(* IEC 61131-3 sources: plcassist-cli/packages/volt-lsp-iec/test-corpus/bakon-nano/Device/Plc Logic/Application/POUs/Calculations (part 4) *)

(* ---- Calc_BottomPos.prg ---- *)
PROGRAM Calc_BottomPos
VAR
END_VAR

//Bereken diepste positie van Z-as (Hoogste) afhankelijk van geselecteerd product plaat.

CASE g_HMI_RCP_Parameters.nProductType  OF
	Prod_Tray_Rectangle_1x1:
		g_sCalculated.rBottomZPos		:= g_HMI_MCH_Parameters.rBottomZPosTrayLarge - g_HMI_RCP_Parameters.rStopHeightKnife;
		g_sCalculated.rAboveProductPos	:= MIN((g_HMI_MCH_Parameters.rBottomZPosTrayLarge - g_HMI_RCP_Parameters.rStartHeightKnife - C_rExtraMarginKnifeHeight),(g_HMI_MCH_Parameters.rBottomZPosTrayLarge - g_HMI_MCH_Parameters.rProdHeightTrayMinimum));
		g_sCalculated.rCrashCheckHeight	:= (g_HMI_MCH_Parameters.rBottomZPosTrayLarge - g_HMI_MCH_Parameters.rProdHeightTrayMinimum + 8); // + 5mm
	Prod_Tray_Rectangle_1x2:
		g_sCalculated.rBottomZPos	:= g_HMI_MCH_Parameters.rBottomZPosTraySmall - g_HMI_RCP_Parameters.rStopHeightKnife;
		g_sCalculated.rAboveProductPos := MIN((g_HMI_MCH_Parameters.rBottomZPosTraySmall - g_HMI_RCP_Parameters.rStartHeightKnife - C_rExtraMarginKnifeHeight),(g_HMI_MCH_Parameters.rBottomZPosTraySmall - g_HMI_MCH_Parameters.rProdHeightTrayMinimum));
		g_sCalculated.rCrashCheckHeight	:= (g_HMI_MCH_Parameters.rBottomZPosTraySmall - g_HMI_MCH_Parameters.rProdHeightTrayMinimum + 8); // + 5mm
	Prod_Tray_Rectangle_2x1:		(* V07.01 *)
		g_sCalculated.rBottomZPos		 := g_HMI_MCH_Parameters.rBottomZPosTrayDouble - g_HMI_RCP_Parameters.rStopHeightKnife;
		g_sCalculated.rAboveProductPos := MIN((g_HMI_MCH_Parameters.rBottomZPosTrayDouble - g_HMI_RCP_Parameters.rStartHeightKnife - C_rExtraMarginKnifeHeight),(g_HMI_MCH_Parameters.rBottomZPosTrayDouble - g_HMI_MCH_Parameters.rProdHeightTrayMinimum));
		g_sCalculated.rCrashCheckHeight	:= (g_HMI_MCH_Parameters.rBottomZPosTrayDouble - g_HMI_MCH_Parameters.rProdHeightTrayMinimum + 8); // + 5mm
	Prod_Tray_Rectangle_1x4:
		g_sCalculated.rBottomZPos	:= g_HMI_MCH_Parameters.rBottomZPosTrayTriple - g_HMI_RCP_Parameters.rStopHeightKnife;
		g_sCalculated.rAboveProductPos := MIN((g_HMI_MCH_Parameters.rBottomZPosTrayTriple - g_HMI_RCP_Parameters.rStartHeightKnife - C_rExtraMarginKnifeHeight),(g_HMI_MCH_Parameters.rBottomZPosTrayTriple - g_HMI_MCH_Parameters.rProdHeightTrayMinimum));
		g_sCalculated.rCrashCheckHeight	:= (g_HMI_MCH_Parameters.rBottomZPosTrayTriple -g_HMI_MCH_Parameters.rProdHeightTrayMinimum + 8); // + 5mm
	Prod_Round_POC_2x1:
		g_sCalculated.rBottomZPos	:= g_HMI_MCH_Parameters.rBottomZPosRound - g_HMI_RCP_Parameters.rStopHeightKnife;
		g_sCalculated.rAboveProductPos := MIN((g_HMI_MCH_Parameters.rBottomZPosRound - g_HMI_RCP_Parameters.rStartHeightKnife - C_rExtraMarginKnifeHeight),(g_HMI_MCH_Parameters.rBottomZPosRound - 10));	(* altijd minimaal 10 mm *)
		g_sCalculated.rCrashCheckHeight	:= (g_HMI_MCH_Parameters.rBottomZPosRound - g_HMI_MCH_Parameters.rProdHeightTrayMinimum + 8); // + 5mm
	Prod_Round_POC_2x2:
		g_sCalculated.rBottomZPos	:= g_HMI_MCH_Parameters.rBottomZPosRoundQuatro - g_HMI_RCP_Parameters.rStopHeightKnife;
		g_sCalculated.rAboveProductPos := MIN((g_HMI_MCH_Parameters.rBottomZPosRoundQuatro - g_HMI_RCP_Parameters.rStartHeightKnife - C_rExtraMarginKnifeHeight),(g_HMI_MCH_Parameters.rBottomZPosRoundQuatro - 10));	(* altijd minimaal 10 mm *)
		g_sCalculated.rCrashCheckHeight	:= (g_HMI_MCH_Parameters.rBottomZPosRoundQuatro - g_HMI_MCH_Parameters.rProdHeightTrayMinimum + 8); // + 5mm
	Prod_Slab_Rectangle_2x1:
		g_sCalculated.rBottomZPos	:= g_HMI_MCH_Parameters.rBottomZPosSlabDouble - g_HMI_RCP_Parameters.rStopHeightKnife;
		g_sCalculated.rAboveProductPos := MIN((g_HMI_MCH_Parameters.rBottomZPosSlabDouble - g_HMI_RCP_Parameters.rStartHeightKnife - C_rExtraMarginKnifeHeight),(g_HMI_MCH_Parameters.rBottomZPosSlab - 10));
		g_sCalculated.rCrashCheckHeight	:= (g_HMI_MCH_Parameters.rBottomZPosSlabDouble - g_HMI_MCH_Parameters.rProdHeightTrayMinimum + 8); // + 5mm
ELSE
		g_sCalculated.rBottomZPos	:= g_HMI_MCH_Parameters.rBottomZPosSlab - g_HMI_RCP_Parameters.rStopHeightKnife;
		g_sCalculated.rAboveProductPos := MIN((g_HMI_MCH_Parameters.rBottomZPosSlab - g_HMI_RCP_Parameters.rStartHeightKnife - C_rExtraMarginKnifeHeight),(g_HMI_MCH_Parameters.rBottomZPosSlab - 10));
		g_sCalculated.rCrashCheckHeight	:= (g_HMI_MCH_Parameters.rBottomZPosSlab - g_HMI_MCH_Parameters.rProdHeightTrayMinimum + 8); // + 5mm
END_CASE

g_sCalculated.rCrashCheckHeight := MIN(g_sCalculated.rCrashCheckHeight, g_sCalculated.rBottomZPos-1);

IF g_HMI_MachCommand.bScanMode THEN
		g_sCalculated.rBottomZPos	:= MIN(g_HMI_MCH_Parameters.rBottomZPosSlab,
										MIN(g_HMI_MCH_Parameters.rBottomZPosSlabDouble,
										MIN(g_HMI_MCH_Parameters.rBottomZPosRoundQuatro,
										MIN(g_HMI_MCH_Parameters.rBottomZPosRound,
										MIN(g_HMI_MCH_Parameters.rBottomZPosTrayDouble,
										MIN(g_HMI_MCH_Parameters.rBottomZPosTrayLarge,
										MIN(g_HMI_MCH_Parameters.rBottomZPosTraySmall,
										g_HMI_MCH_Parameters.rBottomZPosTrayTriple)))))));
		g_sCalculated.rAboveProductPos := 0;
END_IF

g_sCalculated.rAboveProductPos := SEL(g_sMACH.MCL.bActCleaning,g_sCalculated.rAboveProductPos,0); //AC Correctie voor schoonmaak bedrijf waarbij er nog geen bottompos is ingesteld

END_PROGRAM

(* ---- Calc_Init.prg ---- *)
PROGRAM Calc_Init
VAR
	Cnt_pos: INT;
END_VAR

(* Init array *)
FOR Cnt_pos := 1 TO (C_wNumberOfMotionObjects -1)  BY 1 DO
	g_aCuttingPositions[Cnt_pos].X_Target			:=-50;
	g_aCuttingPositions[Cnt_pos].Y_Target			:=-50;
	g_aCuttingPositions[Cnt_pos].A_Target			:=-50;
	g_aCuttingPositions[Cnt_pos].K_Target			:= 0;
	g_aCuttingPositions[Cnt_pos].bPushAwayProduct 	:= FALSE;
	g_aCuttingPositions[Cnt_pos].rPushAwayDistance 	:= 0;
	g_aCuttingPositions[Cnt_pos].bCutPosPossible 	:= TRUE;
	g_aCuttingPositions[Cnt_pos].bCrashDetectCheck 	:= FALSE;
END_FOR

FOR Cnt_pos := 1 TO 100 BY 1 DO
	g_aWastePositions[Cnt_pos].X_Target				:=-50;
	g_aWastePositions[Cnt_pos].Y_Target				:=-50;
	g_aWastePositions[Cnt_pos].A_Target				:=-50;
	g_aWastePositions[Cnt_pos].K_Target				:= 0;
	g_aWastePositions[Cnt_pos].bPushAwayProduct 	:= FALSE;
	g_aWastePositions[Cnt_pos].rPushAwayDistance 	:= 0;
	g_aWastePositions[Cnt_pos].bCutPosPossible 		:= TRUE;
	g_aWastePositions[Cnt_pos].bCrashDetectCheck	:= FALSE;
END_FOR

(*Minimale Afvalrand limieten bepalen*)
CASE G_HMI_RCP_Parameters.nProductType OF
	Prod_Tray_Rectangle_1x2, Prod_Tray_Rectangle_1x1, Prod_Tray_Rectangle_1x4, Prod_Tray_Rectangle_2x1 :	(* Tray products *)
	g_HMI_RCP_Parameters.rSizeTrimRight := MAX( g_HMI_RCP_Parameters.rSizeTrimRight, 0);
	g_HMI_RCP_Parameters.rSizeTrimLeft 	:= MAX( g_HMI_RCP_Parameters.rSizeTrimLeft, 0);
	g_HMI_RCP_Parameters.rSizeTrimFront := MAX( g_HMI_RCP_Parameters.rSizeTrimFront, 0);
	g_HMI_RCP_Parameters.rSizeTrimRear  := MAX( g_HMI_RCP_Parameters.rSizeTrimRear, 0);
END_CASE

(* Determine waste strips front and rear *)
g_bTrimRight		:=	g_HMI_RCP_Parameters.rSizeTrimRight > 0 ;
g_bTrimLeft			:=	g_HMI_RCP_Parameters.rSizeTrimLeft > 0 ;
g_bTrimRear			:=	g_HMI_RCP_Parameters.rSizeTrimFront > 0 ;(*AC 28-11-12: Omgedraaid vanaf HMI INstellingen*)
g_bTrimFront		:=	g_HMI_RCP_Parameters.rSizeTrimRear > 0 ;(*AC 28-11-12: Omgedraaid vanaf HMI INstellingen*)

g_sCuttingPositionsInfo.index := g_sCuttingPositionsInfo.lowerBound;	(* Array counter *)
g_sWastePositionsInfo.index := g_sWastePositionsInfo.lowerBound;

g_sMACH.ERR.bOvershootCorrectionImpossible := FALSE;

END_PROGRAM

(* ---- Calc_Main.prg ---- *)
PROGRAM Calc_Main
VAR

	rCenterPointKnifeInverted: REAL;
	rSizeOfKnife: REAL;
	rCenterPointKnife: REAL;
	n : INT;
	m : INT;
END_VAR

IF g_bCalculationStart AND NOT g_bCalculationDone
THEN
	Calc_Init();

	IF NOT g_HMI_MachCommand.bScanMode THEN

		(* Knife position 90 degrees: (|) *)
		IF NOT Calc_Ver() THEN
			g_sMACH.ERR.bCalcVerError := TRUE;
		END_IF

		IF NOT Calc_Hor() THEN
			g_sMACH.ERR.bCalcHorError := TRUE;
		END_IF

		IF NOT Calc_Dia1_Compact() THEN
			g_sMACH.ERR.bCalcDia1Error := TRUE;
		END_IF

		IF NOT Calc_Dia2_Compact() THEN
			g_sMACH.ERR.bCalcDia2Error := TRUE;
		END_IF

		(*Loopje om afval posities vooraan te zetten*)
		IF g_HMI_RCP_Parameters.bCutWasteFirst AND (g_bTrimFront OR g_bTrimRear OR g_bTrimLeft OR g_bTrimRight) THEN
			FOR n := g_sCuttingPositionsInfo.index + g_sWastePositionsInfo.index  - 2 TO 1 BY -1 DO
				IF n < g_sWastePositionsInfo.index  THEN
					g_aCuttingPositions[n] := g_aWastePositions[n];
				ELSE
					g_aCuttingPositions[n] := g_aCuttingPositions[n - g_sWastePositionsInfo.index +1];
				END_IF
			END_FOR
		END_IF

		(*Loopje voor crash detectie posities*)
		IF gMachConfig.bCrashDetection AND g_HMI_RCP_Parameters.bCutWasteFirst AND
			(g_HMI_RCP_Parameters.nProductType = Prod_Tray_Rectangle_1x1
			OR	g_HMI_RCP_Parameters.nProductType = Prod_Tray_Rectangle_1x2
			OR g_HMI_RCP_Parameters.nProductType = Prod_Tray_Rectangle_1x4
			OR g_HMI_RCP_Parameters.nProductType = Prod_Tray_Rectangle_2x1
			)
		THEN
			m := g_sCuttingPositionsInfo.index + g_sWastePositionsInfo.index  -2 + g_sWastePositionsInfo.index  -1;
			FOR n := g_sCuttingPositionsInfo.index + g_sWastePositionsInfo.index  -2 TO 1 BY -1 DO
				g_aCuttingPositions[m] := g_aCuttingPositions[n];
				m := m -1;
				IF n < g_sWastePositionsInfo.index  THEN
					g_aCuttingPositions[m] := g_aCuttingPositions[n];
					g_aCuttingPositions[m].bPushAwayProduct := FALSE;
					g_aCuttingPositions[m].bCrashDetectCheck := TRUE;
					m := m - 1;
				END_IF
			END_FOR
		END_IF

		(* V13.01, delete all impossible cutting positions *)
		Calc_SkipPositions();
	ELSE
		Calc_Service();
	END_IF

	Calc_BottomPos();	// Calculate Z bottom pos and pos above product

	rSizeOfKnife					:= g_HMI_MCH_Parameters.rSizeOfKnife;
	rCenterPointKnife				:= rSizeOfKnife/2;
	rCenterPointKnifeInverted	:= rSizeOfKnife/2;

	g_rEndTargetX := g_aCuttingPositions[1].X_Target;
	g_rEndTargetY := g_aCuttingPositions[1].Y_Target;
	g_rEndTargetA := g_aCuttingPositions[1].A_Target;
	g_rEndTargetK := g_aCuttingPositions[1].K_Target;
END_IF
g_bCalculationDone := g_bCalculationStart;

END_PROGRAM

(* ---- Calc_Service.prg ---- *)
PROGRAM Calc_Service
VAR
	rStartPointSlab_X: REAL;
	rStartPointSlab_Y: REAL;
	rSizeTrimRear: REAL;
	rSizeTrimRight: REAL;
	nPos: INT;
END_VAR

	nPos	:= 1;

	(* Ronde taart *)
	g_aCuttingPositions[nPos].X_Target := g_HMI_MCH_Parameters.rMidPosRoundCake1_X;
	g_aCuttingPositions[nPos].Y_Target := g_HMI_MCH_Parameters.rMidPosRoundCake1_Y;
	g_aCuttingPositions[nPos].A_Target := 0;
	nPos	:= nPos + 1;

	g_aCuttingPositions[nPos].X_Target := g_HMI_MCH_Parameters.rMidPosRoundCake1_X;
	g_aCuttingPositions[nPos].Y_Target := g_HMI_MCH_Parameters.rMidPosRoundCake1_Y;
	g_aCuttingPositions[nPos].A_Target := 90;
	nPos	:= nPos + 1;

	g_aCuttingPositions[nPos].X_Target := g_HMI_MCH_Parameters.rMidPosRoundCake1_X;
	g_aCuttingPositions[nPos].Y_Target := g_HMI_MCH_Parameters.rMidPosRoundCake1_Y;
	g_aCuttingPositions[nPos].A_Target := 45;
	nPos	:= nPos + 1;

	g_aCuttingPositions[nPos].X_Target := g_HMI_MCH_Parameters.rMidPosRoundCake1_X;
	g_aCuttingPositions[nPos].Y_Target := g_HMI_MCH_Parameters.rMidPosRoundCake1_Y;
	g_aCuttingPositions[nPos].A_Target := 135;
	nPos	:= nPos + 1;

	(* Slab verticaal (|) *)
	rStartPointSlab_X	:= MAX(g_HMI_MCH_Parameters.rStartPointSlab_X, g_HMI_MCH_Parameters.rStartPointTrayLarge_X);
	rStartPointSlab_Y	:= MAX(g_HMI_MCH_Parameters.rStartPointSlab_Y, g_HMI_MCH_Parameters.rStartPointTrayLarge_Y);
	rSizeTrimRight	:= 10;
	rSizeTrimRear		:= 10;

	g_aCuttingPositions[nPos].X_Target := rStartPointSlab_X + rSizeTrimRight;
	g_aCuttingPositions[nPos].Y_Target := rStartPointSlab_Y + rSizeTrimRear + g_HMI_MCH_Parameters.rSizeOfKnife/2;
	g_aCuttingPositions[nPos].A_Target := 90;
	nPos	:= nPos + 1;

	g_aCuttingPositions[nPos].X_Target := rStartPointSlab_X + rSizeTrimRight;
	g_aCuttingPositions[nPos].Y_Target := rStartPointSlab_Y + rSizeTrimRear + g_HMI_MCH_Parameters.rSizeOfKnife / 2 + 65;
	g_aCuttingPositions[nPos].A_Target := 90;
	nPos	:= nPos + 1;

	g_aCuttingPositions[nPos].X_Target := rStartPointSlab_X + rSizeTrimRight + 200;
	g_aCuttingPositions[nPos].Y_Target := rStartPointSlab_Y + rSizeTrimRear + g_HMI_MCH_Parameters.rSizeOfKnife / 2 + 65;
	g_aCuttingPositions[nPos].A_Target := 90;
	nPos	:= nPos + 1;

	g_aCuttingPositions[nPos].X_Target := rStartPointSlab_X + rSizeTrimRight + 200;
	g_aCuttingPositions[nPos].Y_Target := rStartPointSlab_Y + rSizeTrimRear + g_HMI_MCH_Parameters.rSizeOfKnife / 2;
	g_aCuttingPositions[nPos].A_Target := 90;
	nPos	:= nPos + 1;

	g_aCuttingPositions[nPos].X_Target := rStartPointSlab_X + rSizeTrimRight + 400;
	g_aCuttingPositions[nPos].Y_Target := rStartPointSlab_Y + rSizeTrimRear + g_HMI_MCH_Parameters.rSizeOfKnife / 2;
	g_aCuttingPositions[nPos].A_Target := 90;
	nPos	:= nPos + 1;

	g_aCuttingPositions[nPos].X_Target := rStartPointSlab_X + rSizeTrimRight + 400;
	g_aCuttingPositions[nPos].Y_Target := rStartPointSlab_Y + rSizeTrimRear + g_HMI_MCH_Parameters.rSizeOfKnife / 2 + 65;
	g_aCuttingPositions[nPos].A_Target := 90;
	nPos	:= nPos + 1;

	(* Slab horizontal (-----) *)
	g_aCuttingPositions[nPos].X_Target := rStartPointSlab_X + rSizeTrimRight + g_HMI_MCH_Parameters.rSizeOfKnife / 2;
	g_aCuttingPositions[nPos].Y_Target := rStartPointSlab_Y + rSizeTrimRear;
	g_aCuttingPositions[nPos].A_Target := 0;
	nPos	:= nPos + 1;

	g_aCuttingPositions[nPos].X_Target := rStartPointSlab_X + rSizeTrimRight + g_HMI_MCH_Parameters.rSizeOfKnife / 2;
	g_aCuttingPositions[nPos].Y_Target := rStartPointSlab_Y + rSizeTrimRear + 100;
	g_aCuttingPositions[nPos].A_Target := 0;
	nPos	:= nPos + 1;

	g_aCuttingPositions[nPos].X_Target := rStartPointSlab_X + rSizeTrimRight + g_HMI_MCH_Parameters.rSizeOfKnife / 2;
	g_aCuttingPositions[nPos].Y_Target := rStartPointSlab_Y + rSizeTrimRear + 200;
	g_aCuttingPositions[nPos].A_Target := 0;
	nPos	:= nPos + 1;

	g_aCuttingPositions[nPos].X_Target := rStartPointSlab_X + rSizeTrimRight + g_HMI_MCH_Parameters.rSizeOfKnife / 2;
	g_aCuttingPositions[nPos].Y_Target := rStartPointSlab_Y + rSizeTrimRear +300;
	g_aCuttingPositions[nPos].A_Target := 0;
	nPos	:= nPos + 1;

	g_aCuttingPositions[nPos].X_Target := rStartPointSlab_X + rSizeTrimRight + g_HMI_MCH_Parameters.rSizeOfKnife / 2;
	g_aCuttingPositions[nPos].Y_Target := rStartPointSlab_Y + rSizeTrimRear + 400;
	g_aCuttingPositions[nPos].A_Target := 0;
	nPos	:= nPos + 1;

	(* Slab diagonaal, 45 graden, NB: vaste waarden, dus met ander mes kloppen de posities niet!!!! (mes tijdens beurs 315mm) *)
	g_aCuttingPositions[nPos].X_Target := 596; (* 1 *)
	g_aCuttingPositions[nPos].Y_Target := 109;
	g_aCuttingPositions[nPos].A_Target := 45;
	nPos	:= nPos + 1;

	g_aCuttingPositions[nPos].X_Target := 571;
	g_aCuttingPositions[nPos].Y_Target := 134;
	g_aCuttingPositions[nPos].A_Target := 45;
	nPos	:= nPos + 1;

	g_aCuttingPositions[nPos].X_Target := 546;
	g_aCuttingPositions[nPos].Y_Target := 159;
	g_aCuttingPositions[nPos].A_Target := 45;
	nPos	:= nPos + 1;

	g_aCuttingPositions[nPos].X_Target := 521; (* 4 *)
	g_aCuttingPositions[nPos].Y_Target := 184;
	g_aCuttingPositions[nPos].A_Target := 45;
	nPos	:= nPos + 1;

	g_aCuttingPositions[nPos].X_Target := 482.3693;
	g_aCuttingPositions[nPos].Y_Target := 195.3693;
	g_aCuttingPositions[nPos].A_Target := 45;
	nPos	:= nPos + 1;

	g_aCuttingPositions[nPos].X_Target := 509.6307;
	g_aCuttingPositions[nPos].Y_Target := 222.6307;
	g_aCuttingPositions[nPos].A_Target := 45;
	nPos	:= nPos + 1;

	g_aCuttingPositions[nPos].X_Target := 509.6307; (* 7 *)
	g_aCuttingPositions[nPos].Y_Target := 272.6307;
	g_aCuttingPositions[nPos].A_Target := 45;
	nPos	:= nPos + 1;

	g_aCuttingPositions[nPos].X_Target := 432.3693;
	g_aCuttingPositions[nPos].Y_Target := 195.3693;
	g_aCuttingPositions[nPos].A_Target := 45;
	nPos	:= nPos + 1;
	g_aCuttingPositions[nPos].X_Target := 382.3693;
	g_aCuttingPositions[nPos].Y_Target := 195.3693;
	g_aCuttingPositions[nPos].A_Target := 45;
	nPos	:= nPos + 1;

	g_aCuttingPositions[nPos].X_Target := 509.6307; (* 10 *)
	g_aCuttingPositions[nPos].Y_Target := 322.6307;
	g_aCuttingPositions[nPos].A_Target := 45;
	nPos	:= nPos + 1;

END_PROGRAM

(* ---- Calc_SkipPositions.prg ---- *)
PROGRAM Calc_SkipPositions
VAR
	nPosCount : INT;
	nPosCountGood	: INT;
	n					: INT;
END_VAR

(* Delete all impossible cutting positions in array *)

(* init counters *)
nPosCount := 1;
nPosCountGood	:= 1;

(* Do while position in array is a valid calculated value *)
WHILE	((g_aCuttingPositions[nPosCount].X_Target <> -50)
	OR	(g_aCuttingPositions[nPosCount].Y_Target <> -50)
	OR	(g_aCuttingPositions[nPosCount].A_Target <> -50))
	AND nPosCount <= C_wNumberOfMotionObjects
DO
	IF	g_aCuttingPositions[nPosCount].bCutPosPossible THEN
		g_aCuttingPositions[nPosCountGood]	:= g_aCuttingPositions[nPosCount];
		nPosCountGood	:= nPosCountGood + 1;
	END_IF
	nPosCount	:= nPosCount + 1;
END_WHILE

(* Delete unused (double) positions *)
FOR n := nPosCountGood TO nPosCount DO
	IF n <= C_wNumberOfMotionObjects THEN
		g_aCuttingPositions[n].X_Target := -50;
		g_aCuttingPositions[n].Y_Target := -50;
		g_aCuttingPositions[n].A_Target := -50;
	END_IF
END_FOR

g_sMACH.ERR.bMessagePosNotPossible := (nPosCountGood <> nPosCount) AND g_HMI_MCH_Parameters.bSkipImpossiblePositions;

END_PROGRAM
